TYPE ST_CodToNCParam :
STRUCT
	bArrayReseved1: BOOL;     //动子出现标志
	bArrayReseved2: BOOL;     //动子消失标志
	bArrayReseved3: BOOL;
	bArrayReseved4: BOOL;
	bArrayReseved5: BOOL;
	bArrayReseved6: BOOL;
	bArrayReseved7: BOOL;
	bArrayReseved8: BOOL;
	bArrayReseved9: BOOL;
	bArrayReseved10: BOOL;
	bArrayReseved11: BOOL;
	bArrayReseved12: BOOL;
	bArrayReseved13: BOOL;
	bArrayReseved14: BOOL;
	bArrayReseved15: BOOL;
	bArrayReseved16: BOOL;
	nAxisState: UINT;
	nRoadID: UINT;
	fActualPos: LREAL;
	fActualVel: LREAL;
	fActualTorque: LREAL;
END_STRUCT
END_TYPE

(* stored: Version 1.1.0.1, ProductVersion 3.1.4024.12
   DUT ST_CodToNCParam: Id {04c90021-062d-4a00-8d89-2592014acb9b} *)
